Fanuc KAREL source: KT00747.KL

PROGRAM KT00747
%NOLOCKGROUP
VAR
  ARG: ARRAY[4] OF JOINTPOS
  OUT: INTEGER
BEGIN
  OUT = ARRAY_LEN(ARG)
END KT00747
